{attribute 'qualified_only'}
VAR_GLOBAL
	Shutter1OpenRelay : fbMonostableRelay;
	Shutter1CloseRelay : fbMonostableRelay;
END_VAR

(* stored: Version 1.1.0.1
   GVL gvlRelays: Id {b5dc0003-b812-4326-a60f-582349aca143} *)
